{region 'Documentation'}
(*!
<summary>Checks whether the LINT value is inside the inclusive range.</summary>
<description>

Minimum &gt; Maximum reports Error during active evaluation; equal bounds are
valid.

</description>
*)
{endregion}
FUNCTION_BLOCK AssertInRange_LInt EXTENDS AssertionBase
VAR_INPUT
    IN : LINT; //! Actual value checked or observed by this Assertion.
    Minimum : LINT; //! Inclusive lower bound of the comparison; for a range, must not exceed Maximum.
    Maximum : LINT; //! Inclusive upper bound of the comparison; for a range, must not be below Minimum.
END_VAR

SUPER^();

{region 'Documentation'}
(*!
<summary>Check whether the LINT value is inside the inclusive range.</summary>
*)
{endregion}
METHOD PROTECTED Assert
VAR
    Message : STRING(GVL_Constants.MessageLength);
    MinimumText : STRING(GVL_Constants.AssertionValueLength);
    MaximumText : STRING(GVL_Constants.AssertionValueLength);
    ActualText : STRING(GVL_Constants.AssertionValueLength);
END_VAR
IF NOT EvaluationActive THEN
    RETURN;
END_IF;

IF Result = E_Result.Error THEN
    RETURN;
END_IF;

IF Minimum > Maximum THEN
    MinimumText := LINT_TO_STRING(Minimum);
    MaximumText := LINT_TO_STRING(Maximum);
    Message := CONCAT('Assertion error: minimum exceeds maximum. Minimum = ',
        MinimumText);
    Message := CONCAT(Message, ', Maximum = ');
    Message := CONCAT(Message, MaximumText);
    Message := CONCAT(Message, '.');
    Error(Message := Message);
    RETURN;
END_IF;

IF Result = E_Result.Failed THEN
    RETURN;
END_IF;

IF (IN < Minimum) OR (IN > Maximum) THEN
    MinimumText := LINT_TO_STRING(Minimum);
    MaximumText := LINT_TO_STRING(Maximum);
    ActualText := LINT_TO_STRING(IN);
    Message := CONCAT('Assertion failed: value is outside allowed range. Minimum = ',
        MinimumText);
    Message := CONCAT(Message, ', Maximum = ');
    Message := CONCAT(Message, MaximumText);
    Message := CONCAT(Message, ', Actual = ');
    Message := CONCAT(Message, ActualText);
    Message := CONCAT(Message, '.');
    Fail(Message := Message);
    RETURN;
END_IF;

Pass();
END_METHOD

END_FUNCTION_BLOCK

(* stored: Version 1.1.0.1
   POU AssertInRange_LInt: Id {1a2d3275-f7f1-403f-851a-2bfde37af8ae}, SpecialFunc None
   Folder Internal: Id {9b39e530-68a3-4fcd-8876-ffd99e872fcd}
   Method Assert: Id {bad169d3-b79a-4fdd-8ecf-440e46b1809d} *)
